Staubli VAL3: main.pgx

public program main()
  local pointRx l_pPoint
  local num l_nResult
  local tool l_tTool
begin
  //  nLastLib=-1
  do
//    call saveData:getTool(saveData:nJogTool,l_tTool)
//    l_pPoint=here(l_tTool,world)

    call areaCheck()
    call checkPoint()


    delay(0)
  until false

end
